(* IEC 61131-3 sources: Caravan/Stations/MachineControl/MachineControl/Network/Heizung_NET, 2 files *)

(* ---- ONE_Heizung_NET_Table-TAB-EPM-01.st ---- *)
#define OBJECTS_CONFIG

FUNCTION GLOBAL TAB ONE_Heizung_NET
-1$UINT, 0$UINT,
0$UINT, 0$UINT,

1$UDINT,
TO_UDINT(3440325224), "TempControl_Class", 0$UINT, 0$UINT, 1$UINT,

_NO_ATTR, TO_UDINT(3229092335), "TEMPCONTROL_CLASS1",

//Internal connections
0$UDINT,
0$UDINT,
0$UDINT,
0$UDINT,

//Initialization values
0$UDINT,
1$UDINT,
TO_UDINT(0), "TempHZS_C", TO_UDINT(0),//|Heizung_NET.TempControl_Class1.TempHZS_C;

//Symbolic initialization values
0$UDINT,
0$UDINT,

//Initialization of string values
0$UDINT,
0$UDINT,

//Configuration of tasks (RealTime, Cyclic, Background)
0$UDINT,
0$UDINT,

0$UDINT,
1$UDINT,
TO_UDINT(0), (50)$UDINT, 4194303$DINT, 	//TEMPCONTROL_CLASS1

0$UDINT,
0$UDINT,

//External connections
0$UDINT,
6$UDINT,
TO_UDINT(0), "TempHZS_C", C_DIR, TO_UDINT(1518191916), "LseEasy","ActTemperature",
TO_UDINT(0), "ActualRoomTemp_C", C_DIR, TO_UDINT(3157766682), "AI0881","TMP_3",
TO_UDINT(0), "ActualUltraheatTemp_C", C_DIR, TO_UDINT(3157766682), "AI0881","TMP_4",
TO_UDINT(0), "SetFanSpeed_C", C_DIR, TO_UDINT(542619847), "SR0201","SetSpeed",
TO_UDINT(0), "MotorRunStop_C", C_DIR, TO_UDINT(542619847), "SR0201","Enable",
TO_UDINT(0), "HeaterRun_C", C_DIR, TO_UDINT(59516340), "TO1611","Output2",

//Magic internal connections
0$UDINT,
0$UDINT,

//Configuration of timeslots of tasks (RealTime, Cyclic)
#ifdef __LSLLDR_TIMESLOTS__
0$UDINT,
0$UDINT,

0$UDINT,
0$UDINT,

#endif //__LSLLDR_TIMESLOTS__

//MultiMaster connections
#ifdef __LSLLDR_MULTIMASTER__
0$UDINT,
0$UDINT,
#endif //__LSLLDR_MULTIMASTER__

//Configuration for task ID (RealTime, CyclicTime)
#ifdef __LSLLDR_TASKID__
"\\\\TASKS2  "
0$UDINT,
0$UDINT,

0$UDINT,
1$UDINT,
(0)$UDINT, 	//TEMPCONTROL_CLASS1

0$UDINT,
0$UDINT,

#endif //__LSLLDR_TASKID__

END_FUNCTION

(* ---- ONE_Heizung_NET_Table.st ---- *)
#define OBJECTS_CONFIG

FUNCTION GLOBAL TAB ONE_Heizung_NET
-1$UINT, 0$UINT,
0$UINT, 0$UINT,

2$UDINT,
TO_UDINT(1724373636), "DayNightSplitter_Class", 0$UINT, 0$UINT, 1$UINT,
TO_UDINT(3440325224), "TempControl_Class", 0$UINT, 0$UINT, 1$UINT,

_NO_ATTR, TO_UDINT(1768910676), "DAYNIGHTSPLITTER_CLASS1",

_NO_ATTR, TO_UDINT(3229092335), "TEMPCONTROL_CLASS1",

//Internal connections
0$UDINT,
0$UDINT,
0$UDINT,
5$UDINT,
TO_UDINT(0), "DesiredHZSTemp", TO_UDINT(1), "SetTempHZS_s",
TO_UDINT(0), "DesiredRoomTemp", TO_UDINT(1), "SetRoomTemp_S",
TO_UDINT(0), "DesiredHeaterPWR", TO_UDINT(1), "HeaterOn_S",
TO_UDINT(0), "DesiredFanMode", TO_UDINT(1), "FanMode_S",
TO_UDINT(0), "DesiredFanSpeed", TO_UDINT(1), "FanSpeed_S",

//Initialization values
0$UDINT,
2$UDINT,
TO_UDINT(1), "TempHZS_C", TO_UDINT(0),//|Heizung_NET.TempControl_Class1.TempHZS_C;
TO_UDINT(1), "ActualUltraheatTemp_C", TO_UDINT(0),//|Heizung_NET.TempControl_Class1.ActualUltraheatTemp_C;

//Symbolic initialization values
0$UDINT,
0$UDINT,

//Initialization of string values
0$UDINT,
0$UDINT,

//Configuration of tasks (RealTime, Cyclic, Background)
0$UDINT,
0$UDINT,

0$UDINT,
2$UDINT,
TO_UDINT(0), (-2147483448)$UDINT, 4194303$DINT, 	//DAYNIGHTSPLITTER_CLASS1
TO_UDINT(1), (50)$UDINT, 4194303$DINT, 	//TEMPCONTROL_CLASS1

0$UDINT,
0$UDINT,

//External connections
0$UDINT,
9$UDINT,
TO_UDINT(0), "OC_ToTimerClass", C_DIR, TO_UDINT(1302809437), "Timer_Class1","ClassSvr",
TO_UDINT(1), "TempHZS_C", C_DIR, TO_UDINT(1518191916), "LseEasy","ActTemperature",
TO_UDINT(1), "ActualRoomTemp_C", C_DIR, TO_UDINT(3157766682), "AI0881","TMP_3",
TO_UDINT(1), "ActualUltraheatTemp_C", C_DIR, TO_UDINT(3157766682), "AI0881","TMP_4",
TO_UDINT(1), "SetFanSpeed_C", C_DIR, TO_UDINT(542619847), "SR0201","SetSpeed",
TO_UDINT(1), "MotorRunStop_C", C_DIR, TO_UDINT(542619847), "SR0201","Enable",
TO_UDINT(1), "HeaterRun_C", C_DIR, TO_UDINT(59516340), "TO1611","Output2",
TO_UDINT(1), "HeaterOn_C", C_DIR, TO_UDINT(59516340), "TO1611","Output1",
TO_UDINT(1), "Heater200Watt_C", C_DIR, TO_UDINT(59516340), "TO1611","Output3",

//Magic internal connections
0$UDINT,
0$UDINT,

//Configuration of timeslots of tasks (RealTime, Cyclic)
#ifdef __LSLLDR_TIMESLOTS__
0$UDINT,
0$UDINT,

0$UDINT,
0$UDINT,

#endif //__LSLLDR_TIMESLOTS__

//MultiMaster connections
#ifdef __LSLLDR_MULTIMASTER__
0$UDINT,
0$UDINT,
#endif //__LSLLDR_MULTIMASTER__

//Configuration for task ID (RealTime, CyclicTime)
#ifdef __LSLLDR_TASKID__
"\\\\TASKS2  "
0$UDINT,
0$UDINT,

0$UDINT,
2$UDINT,
(0)$UDINT, 	//DAYNIGHTSPLITTER_CLASS1
(0)$UDINT, 	//TEMPCONTROL_CLASS1

0$UDINT,
0$UDINT,

#endif //__LSLLDR_TASKID__

END_FUNCTION
